(* IEC 61131-3 sources: llm-plc-st-eval/data/calibracion/gemini-3.1-pro-preview/B1/zero_shot, 3 files *)

(* ---- ejec_1.st ---- *)
```iecst
FUNCTION_BLOCK FB_Motor
VAR_INPUT
    btnMarcha : BOOL; // TRUE al pulsar (Contacto NA)
    btnParo   : BOOL; // TRUE al pulsar (Asumiendo lógica positiva para el ejemplo)
    btnEmerg  : BOOL; // TRUE al pulsar (Asumiendo lógica positiva para el ejemplo)
END_VAR

VAR_OUTPUT
    motorOn   : BOOL; // TRUE = Motor encendido, FALSE = Motor detenido
END_VAR

VAR
    rtMarcha  : R_TRIG; // Detector de flanco ascendente para el botón de marcha
END_VAR

// 1. Detectar el flanco ascendente (transición de FALSE a TRUE) del botón de marcha.
// Esto evita el rearranque automático si el botón se mantiene pulsado tras una emergencia.
rtMarcha(CLK := btnMarcha);

// 2. Lógica de control del motor (Enclavamiento con prioridad al paro).
// El motor se enciende con el flanco de marcha o se mantiene encendido (motorOn),
// siempre y cuando no se pulse el paro normal ni el paro de emergencia.
motorOn := (motorOn OR rtMarcha.Q) AND NOT btnParo AND NOT btnEmerg;

END_FUNCTION_BLOCK
```

(* ---- ejec_2.st ---- *)
```iecst
FUNCTION_BLOCK FB_Motor
VAR_INPUT
    btnMarcha : BOOL; // TRUE al pulsar (arranque)
    btnParo   : BOOL; // TRUE al pulsar (parada normal)
    btnEmerg  : BOOL; // TRUE al pulsar (parada de emergencia)
END_VAR

VAR_OUTPUT
    motorOn   : BOOL; // TRUE = Motor en marcha, FALSE = Motor detenido
END_VAR

VAR
    trigMarcha : R_TRIG; // Detección de flanco para evitar rearranque automático
END_VAR

// Detectar flanco ascendente del botón de marcha
trigMarcha(CLK := btnMarcha);

// Lógica de control: Prioridad a la parada
IF btnEmerg OR btnParo THEN
    motorOn := FALSE;
// Arranque por flanco para exigir soltar y volver a pulsar tras una emergencia
ELSIF trigMarcha.Q THEN
    motorOn := TRUE;
END_IF;

END_FUNCTION_BLOCK
```

(* ---- ejec_3.st ---- *)
```iecst
FUNCTION_BLOCK FB_Motor
VAR_INPUT
    btnMarcha : BOOL; // Botón de marcha (arranque)
    btnParo   : BOOL; // Botón de paro normal (TRUE = pulsado para detener)
    btnEmerg  : BOOL; // Botón de paro de emergencia (TRUE = pulsado para detener)
END_VAR

VAR_OUTPUT
    motorOn   : BOOL; // Señal de activación del motor
END_VAR

VAR
    flancoMarcha : R_TRIG; // Detector de flanco ascendente estándar IEC 61131-3
END_VAR

// Detectar el flanco positivo (pulsación) del botón de marcha.
// Esto evita el rearranque automático si el botón se mantiene pulsado tras una emergencia.
flancoMarcha(CLK := btnMarcha);

// Lógica de control del motor (Enclavamiento)
// Prioridad a las señales de paro (NOT btnParo AND NOT btnEmerg)
motorOn := (flancoMarcha.Q OR motorOn) AND NOT btnParo AND NOT btnEmerg;

END_FUNCTION_BLOCK
```
